(* IEC 61131-3 sources: GenAI/codesys_service/demo, 4 files *)

(* ---- stdlib_strings.st ---- *)
FUNCTION_BLOCK StdlibStrings
VAR_INPUT
    textA : STRING(80) := 'Hello';
    textB : STRING(80) := 'World';
END_VAR
VAR_OUTPUT
    n : INT;
    midOut : STRING(80);
    leftOut : STRING(80);
    rightOut : STRING(80);
    concatOut : STRING(80);
    insertOut : STRING(80);
    deleteOut : STRING(80);
    replaceOut : STRING(80);
    findPos : INT;
END_VAR

(* Minimal regression for the CODESYS Standard Library string functions. *)
n := LEN(textA);
midOut := MID(textA, 2, 2);
leftOut := LEFT(textA, 3);
rightOut := RIGHT(textA, 3);
concatOut := CONCAT(textA, textB);
insertOut := INSERT(textA, 'XY', 2);
deleteOut := DELETE(textA, 2, 2);
replaceOut := REPLACE(textA, 'XY', 2, 2);
findPos := FIND(textA, 'llo');

(* ---- motor_start_stop.bad.st ---- *)
(* 故意写坏的一段 ST，用于验证静态检查能不能挡住低级错误。
   预期：E001（IF 未闭合）+ E004（= 当赋值用）+ W101（Motor2 未声明）+ W102（缺分号） *)
PROGRAM PLC_PRG_BAD
VAR
    StartBtn : BOOL;
    StopBtn  : BOOL;
    Motor    : BOOL;
END_VAR

IF StartBtn AND NOT StopBtn THEN
    Motor = TRUE
    Motor2 := TRUE;

(* ---- motor_start_stop.logicbug.st ---- *)
(* 逻辑有缺陷的版本：只处理了停止按钮，漏了急停 EStop。
   预期：TC01 通过，TC03 失败（急停不能停机）。 *)
PROGRAM PLC_PRG
VAR
    StartBtn : BOOL;
    StopBtn  : BOOL;
    EStop    : BOOL;
    Motor    : BOOL;
END_VAR

IF StartBtn AND NOT StopBtn THEN
    Motor := TRUE;
END_IF;

IF StopBtn THEN
    Motor := FALSE;
END_IF;

(* ---- motor_start_stop.st ---- *)
(* ============================================================
   示例：电机启停控制（对应大作业第六章示例题）
   文件约定：包含 POU 头 + VAR 声明 + 实现体，
   结尾不写 END_PROGRAM（CODESYS 文本化 POU 中它是隐含的）。
   ============================================================ *)
PROGRAM PLC_PRG
VAR
    StartBtn : BOOL;   (* 启动按钮 *)
    StopBtn  : BOOL;   (* 停止按钮 *)
    EStop    : BOOL;   (* 急停信号 *)
    Motor    : BOOL;   (* 电机运行输出 *)
END_VAR

(* 停止/急停优先级高于启动；启动按钮松开后由 Motor 自保持 *)
IF (StopBtn OR EStop) THEN
    Motor := FALSE;
ELSIF (StartBtn AND NOT StopBtn AND NOT EStop) THEN
    Motor := TRUE;
END_IF;
